PROGRAM Main
VAR
	nSeed : ULINT := 0;
	fbTickCounter : FB_TickCounter;
	bAutoMode : BOOL := FALSE;
	nAutoTickInterval : UDINT := 50;
	
	fbTypeTest : FB_TypeTest(nSeed := nSeed);
	fbStringTest : FB_StringTest(nSeed := nSeed);
	fbStructTest : FB_StructPackingTest(nSeed := nSeed);
	fbEnumTest : FB_EnumTest(nSeed := nSeed);
	fbBitPackingTest : FB_BitPackingTest(nSeed := nSeed);
	fbArrayTest : FB_ArrayTest(nSeed := nSeed);
	fbWriteTest : FB_WriteTest;
	
	fbGvlTest : FB_GvlTest(nSeed := nSeed);
	
	{attribute 'some_made_up_var_key':='some_made_up_var_value'}
	fbAttributeTest : FB_AttributeTest;	
END_VAR

fbTypeTest();
fbStringTest();
fbStructTest();
fbEnumTest();
fbBitPackingTest();
fbArrayTest();
fbWriteTest();

fbGvlTest();

fbAttributeTest();

fbTickCounter(bExecute := bAutoMode, nAutoTickInterval := nAutoTickInterval);

IF bAutoMode AND fbTickCounter.bTrigger THEN
	nSeed := nSeed + 1;
END_IF

END_PROGRAM

(* stored: Version 1.1.0.1, ProductVersion 3.1.4026.19
   POU Main: Id {151bda18-a213-42d0-86e0-e79837f085e9}, SpecialFunc None *)
